(* Logix 5000 project; controller R400_500_XLS vendor 1 type 14 code 216 rev 31.11; software revision 31.01; part 17 of 32 *)
(* tags used below, declared in another part *)
   bResetAllCycle : BOOL;
   Calib : SINT;
   CalibCnt : SINT;   // Calibration Step Counter
   CalibData : UDT_SCALE[8];
   CalibEnabled : BOOL;   // RTD Calibration Enabled bit
   CalibIndex : DINT;   // Calibration Pointer
   CustomCycleIterator : DINT;
   CycleDryingStandard : UDT_DRY;
   CycleModifBuffer : UDT_CYCLE;
   Cycles : UDT_CYCLE[11];
   CyclesDefault : UDT_CYCLE[7];   // Preliminary Data block to reset Cycles Values
   CycleSmartDryingHeatSens : UDT_DRY;
   CycleSmartDryingRegular : UDT_DRY;
   CycleWith_NonRecircFRinseDefault : UDT_FRINSE;
   CycleWith_RecircFRinseDefault : UDT_FRINSE;
   CycleWithoutDry : UDT_DRY;
   CycleWithoutFRinseWithoutTankDefault : UDT_FRINSE;
   CycleWithoutFRinseWithTankDefault : UDT_FRINSE;
   DESCALER : SINT;
   DRYING : DINT;   // Drying id number
   ENVIRO_CARE : SINT;
   EXTRA_CARE : SINT;
   FC83_AutoSpeed : BOOL;   // Cycle pump speed selection
   FC83_AutoWtrLevel : BOOL;   // Cycle water level selection
   FC83_CyclePerm : BOOL;   // Cycle permission selection
   M : DINT[5];   // Memory Bits
   ONS_FC84 : SINT;
   PLASTIC_CARE : SINT;
   ResetCycleName : BOOL;
   RINSE_CARE : SINT;
   Run : DINT;
   STANDARD : SINT;
   Supervisor : DINT;
   USER_DEFINED_11 : SINT;
   USER_DEFINED_7 : SINT;
   CycleName : STRING[12];
   CycleNameDefault : STRING[12];
   CyclePtr : DINT;   // Cycle Pointeur
   DryTemp : REAL;
   I_Dry_RTD : DINT;   // Drying RTD
   I_Pw_Tnk_RTD : DINT;   // Pure water tank RTD
   I_Smp_RTD : DINT;   // Sump RTD
   NumInput : UDT_NUMERIC_INPUT[65];   // Numeric input
   PureWaterTankTemp : REAL;   // Pure water tank temperature
   Screen_Ctrl : DINT;   // PLC Screen Request
   StringInput : UDT_STRING_INPUT[6];
   SumpTemp : REAL;   // Sump temperature in °C
   Tpb : DINT[11];
   TpbImage : DINT[11];
   Unit : Hrdwre;   // Unit Configuration
(* MainProgram, continued *)

ROUTINE SPV_4_CycleNames   (* ladder *)
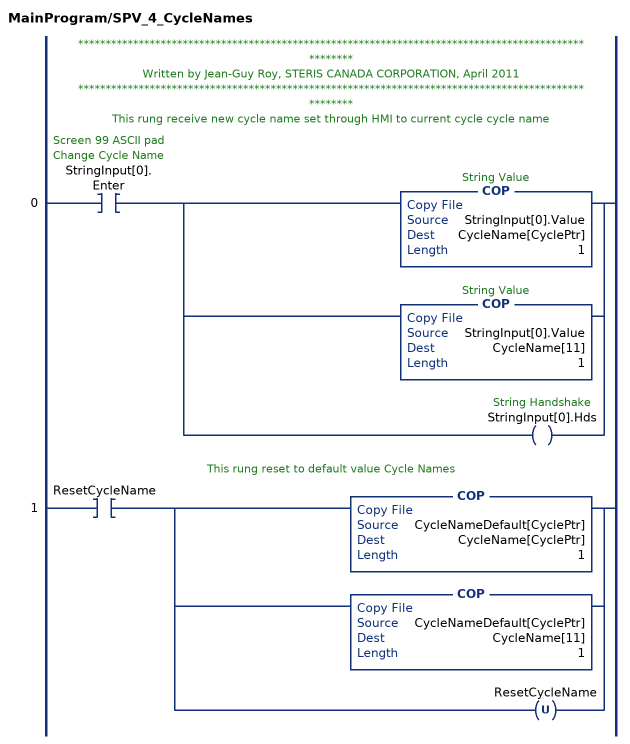
   // ****************************************************************************************************
   // Written by Jean-Guy Roy, STERIS CANADA CORPORATION, April 2011
   // ****************************************************************************************************
   // This rung receive new cycle name set through HMI to current cycle cycle name
   0: XIC(StringInput[0].Enter)[COP(StringInput[0].Value,CycleName[CyclePtr],1) ,COP(StringInput[0].Value,CycleName[11],1) ,OTE(StringInput[0].Hds) ];
   // This rung reset to default value Cycle Names
   1: XIC(ResetCycleName)[COP(CycleNameDefault[CyclePtr],CycleName[CyclePtr],1) ,COP(CycleNameDefault[CyclePtr],CycleName[11],1) ,OTU(ResetCycleName) ];
END_ROUTINE

ROUTINE SPV_8_ResetToDefaultCyclesValues   (* ladder *)
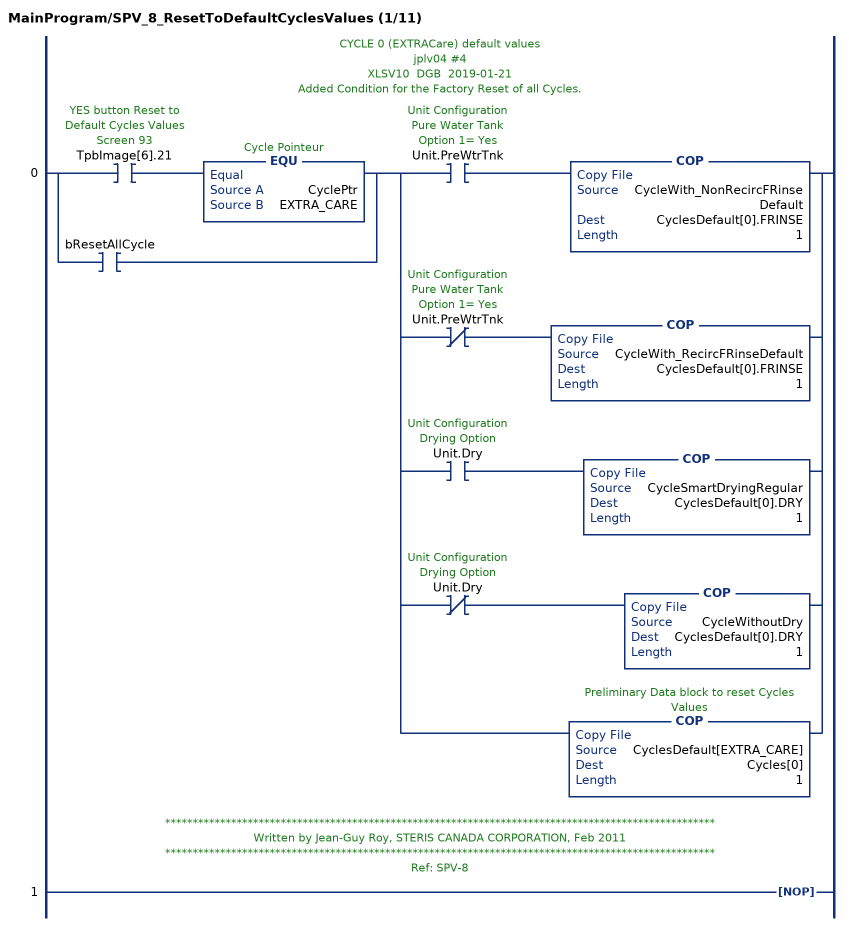
   // CYCLE 0 (EXTRACare) default values
   // jplv04 #4
   // XLSV10  DGB  2019-01-21
   // Added Condition for the Factory Reset of all Cycles.
   0: [XIC(TpbImage[6].21) EQU(CyclePtr,EXTRA_CARE) ,XIC(bResetAllCycle) ][XIC(Unit.PreWtrTnk) COP(CycleWith_NonRecircFRinseDefault,CyclesDefault[0].FRINSE,1) ,XIO(Unit.PreWtrTnk) COP(CycleWith_RecircFRinseDefault,CyclesDefault[0].FRINSE,1) ,XIC(Unit.Dry) COP(CycleSmartDryingRegular,CyclesDefault[0].DRY,1) ,XIO(Unit.Dry) COP(CycleWithoutDry,CyclesDefault[0].DRY,1) ,COP(CyclesDefault[EXTRA_CARE],Cycles[0],1) ];
   // ****************************************************************************************************
   // Written by Jean-Guy Roy, STERIS CANADA CORPORATION, Feb 2011
   // ****************************************************************************************************
   // Ref: SPV-8
   1: NOP();
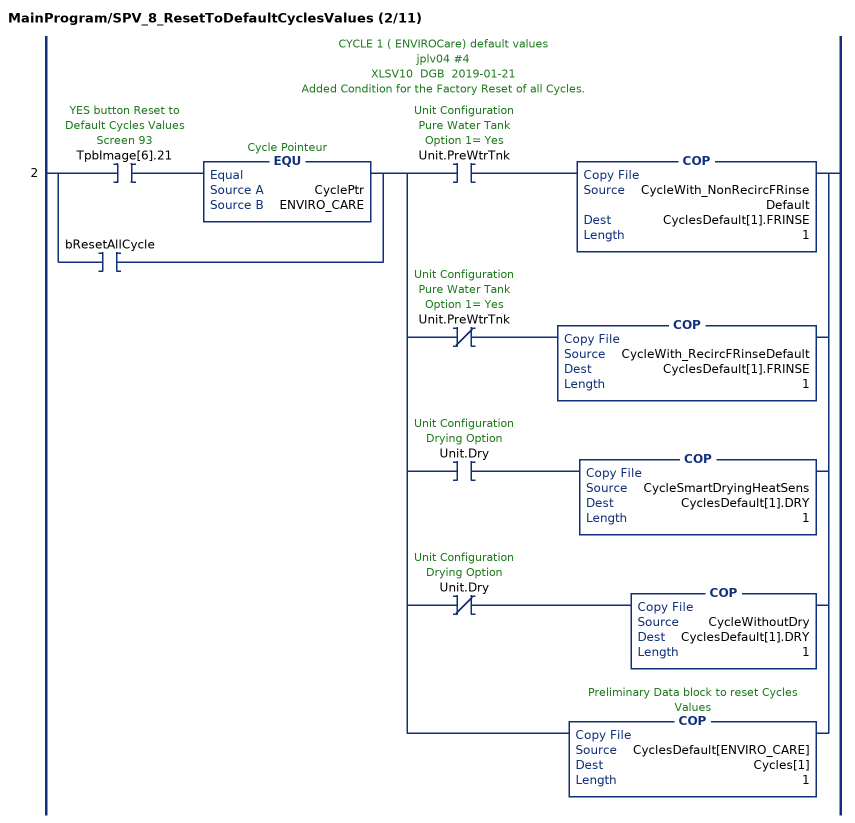
   // CYCLE 1 ( ENVIROCare) default values
   // jplv04 #4
   // XLSV10  DGB  2019-01-21
   // Added Condition for the Factory Reset of all Cycles.
   2: [XIC(TpbImage[6].21) EQU(CyclePtr,ENVIRO_CARE) ,XIC(bResetAllCycle) ][XIC(Unit.PreWtrTnk) COP(CycleWith_NonRecircFRinseDefault,CyclesDefault[1].FRINSE,1) ,XIO(Unit.PreWtrTnk) COP(CycleWith_RecircFRinseDefault,CyclesDefault[1].FRINSE,1) ,XIC(Unit.Dry) COP(CycleSmartDryingHeatSens,CyclesDefault[1].DRY,1) ,XIO(Unit.Dry) COP(CycleWithoutDry,CyclesDefault[1].DRY,1) ,COP(CyclesDefault[ENVIRO_CARE],Cycles[1],1) ];
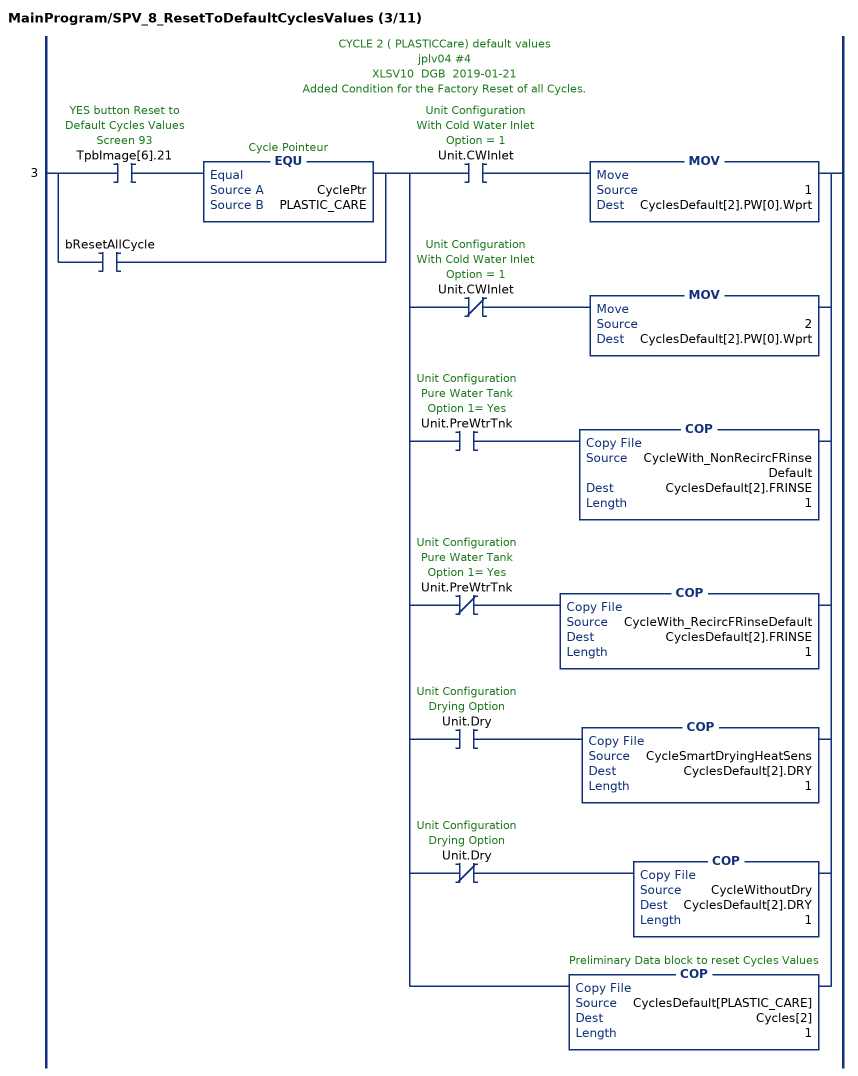
   // CYCLE 2 ( PLASTICCare) default values
   // jplv04 #4
   // XLSV10  DGB  2019-01-21
   // Added Condition for the Factory Reset of all Cycles.
   3: [XIC(TpbImage[6].21) EQU(CyclePtr,PLASTIC_CARE) ,XIC(bResetAllCycle) ][XIC(Unit.CWInlet) MOV(1,CyclesDefault[2].PW[0].Wprt) ,XIO(Unit.CWInlet) MOV(2,CyclesDefault[2].PW[0].Wprt) ,XIC(Unit.PreWtrTnk) COP(CycleWith_NonRecircFRinseDefault,CyclesDefault[2].FRINSE,1) ,XIO(Unit.PreWtrTnk) COP(CycleWith_RecircFRinseDefault,CyclesDefault[2].FRINSE,1) ,XIC(Unit.Dry) COP(CycleSmartDryingHeatSens,CyclesDefault[2].DRY,1) ,XIO(Unit.Dry) COP(CycleWithoutDry,CyclesDefault[2].DRY,1) ,COP(CyclesDefault[PLASTIC_CARE],Cycles[2],1) ];
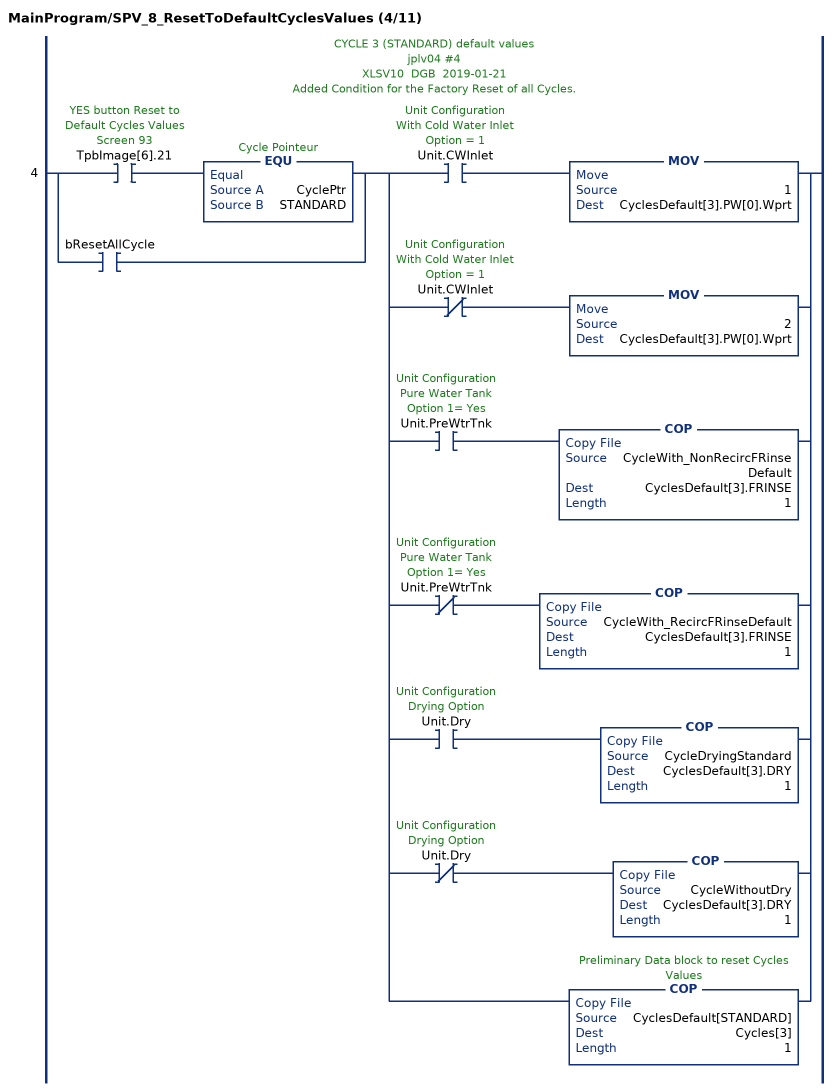
   // CYCLE 3 (STANDARD) default values
   // jplv04 #4
   // XLSV10  DGB  2019-01-21
   // Added Condition for the Factory Reset of all Cycles.
   4: [XIC(TpbImage[6].21) EQU(CyclePtr,STANDARD) ,XIC(bResetAllCycle) ][XIC(Unit.CWInlet) MOV(1,CyclesDefault[3].PW[0].Wprt) ,XIO(Unit.CWInlet) MOV(2,CyclesDefault[3].PW[0].Wprt) ,XIC(Unit.PreWtrTnk) COP(CycleWith_NonRecircFRinseDefault,CyclesDefault[3].FRINSE,1) ,XIO(Unit.PreWtrTnk) COP(CycleWith_RecircFRinseDefault,CyclesDefault[3].FRINSE,1) ,XIC(Unit.Dry) COP(CycleDryingStandard,CyclesDefault[3].DRY,1) ,XIO(Unit.Dry) COP(CycleWithoutDry,CyclesDefault[3].DRY,1) ,COP(CyclesDefault[STANDARD],Cycles[3],1) ];
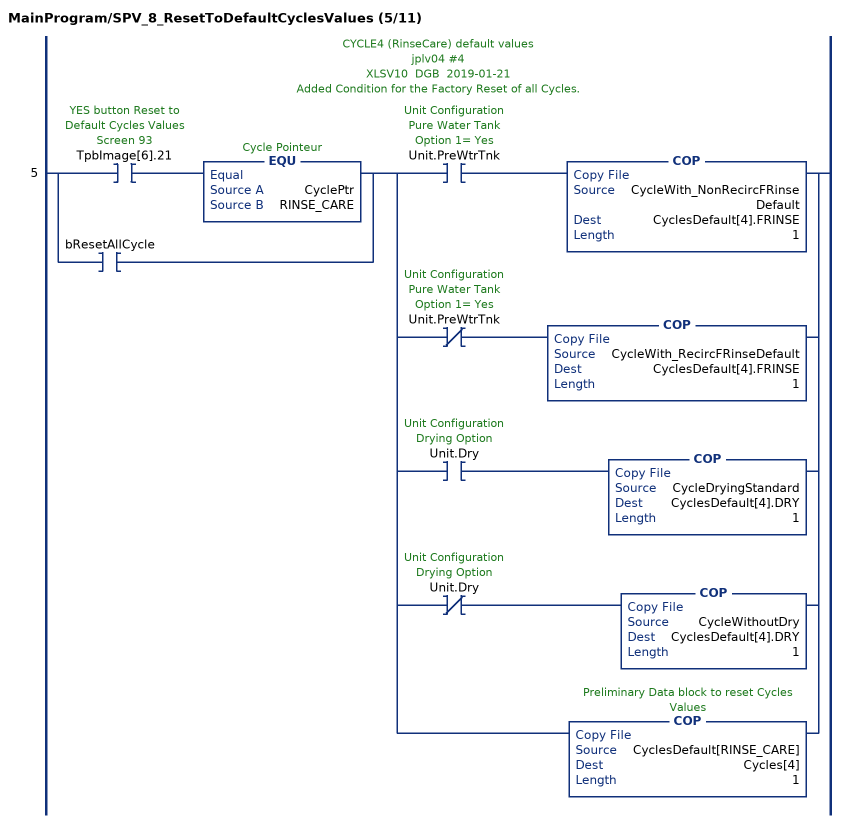
   // CYCLE4 (RinseCare) default values
   // jplv04 #4
   // XLSV10  DGB  2019-01-21
   // Added Condition for the Factory Reset of all Cycles.
   5: [XIC(TpbImage[6].21) EQU(CyclePtr,RINSE_CARE) ,XIC(bResetAllCycle) ][XIC(Unit.PreWtrTnk) COP(CycleWith_NonRecircFRinseDefault,CyclesDefault[4].FRINSE,1) ,XIO(Unit.PreWtrTnk) COP(CycleWith_RecircFRinseDefault,CyclesDefault[4].FRINSE,1) ,XIC(Unit.Dry) COP(CycleDryingStandard,CyclesDefault[4].DRY,1) ,XIO(Unit.Dry) COP(CycleWithoutDry,CyclesDefault[4].DRY,1) ,COP(CyclesDefault[RINSE_CARE],Cycles[4],1) ];
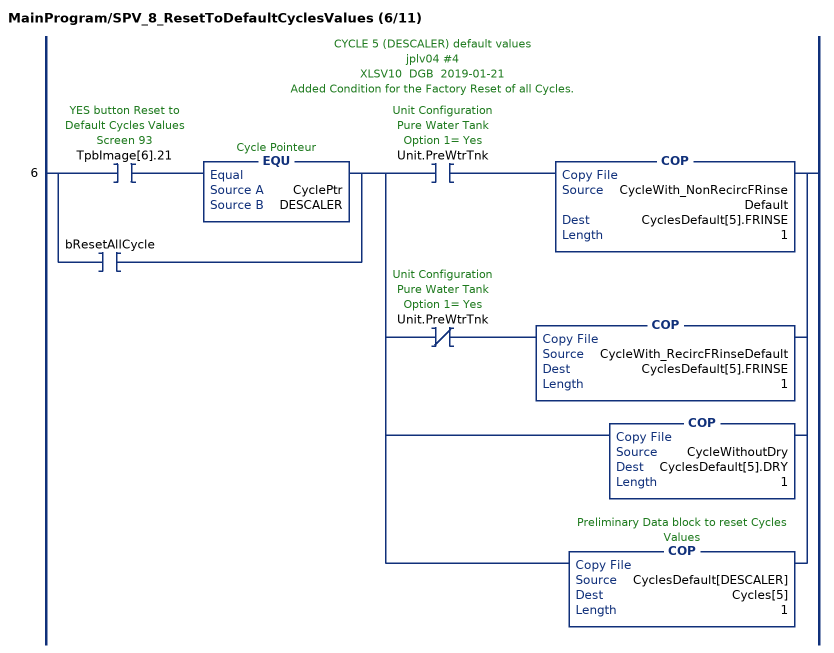
   // CYCLE 5 (DESCALER) default values
   // jplv04 #4
   // XLSV10  DGB  2019-01-21
   // Added Condition for the Factory Reset of all Cycles.
   6: [XIC(TpbImage[6].21) EQU(CyclePtr,DESCALER) ,XIC(bResetAllCycle) ][XIC(Unit.PreWtrTnk) COP(CycleWith_NonRecircFRinseDefault,CyclesDefault[5].FRINSE,1) ,XIO(Unit.PreWtrTnk) COP(CycleWith_RecircFRinseDefault,CyclesDefault[5].FRINSE,1) ,COP(CycleWithoutDry,CyclesDefault[5].DRY,1) ,COP(CyclesDefault[DESCALER],Cycles[5],1) ];
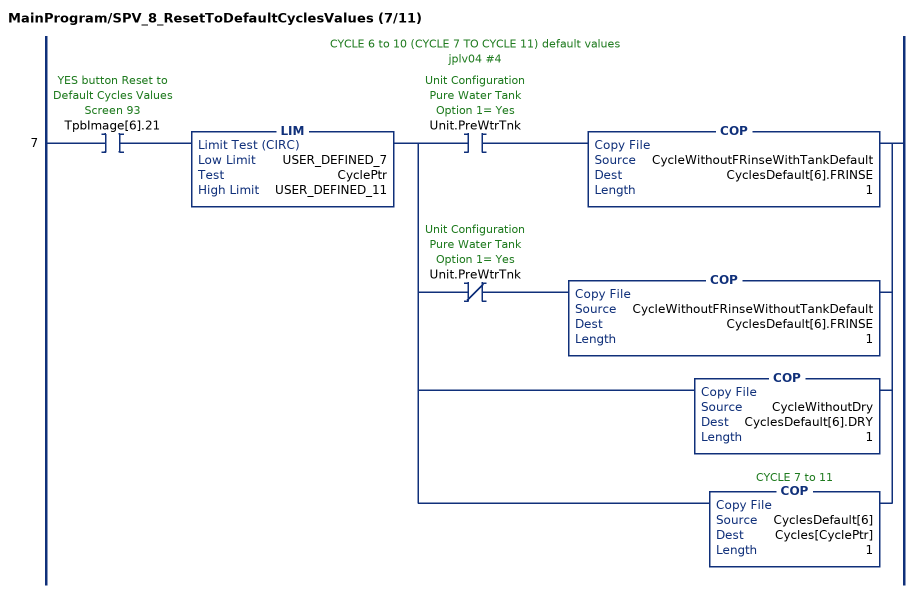
   // CYCLE 6 to 10 (CYCLE 7 TO CYCLE 11) default values
   // jplv04 #4
   7: XIC(TpbImage[6].21)LIM(USER_DEFINED_7,CyclePtr,USER_DEFINED_11)[XIC(Unit.PreWtrTnk) COP(CycleWithoutFRinseWithTankDefault,CyclesDefault[6].FRINSE,1) ,XIO(Unit.PreWtrTnk) COP(CycleWithoutFRinseWithoutTankDefault,CyclesDefault[6].FRINSE,1) ,COP(CycleWithoutDry,CyclesDefault[6].DRY,1) ,COP(CyclesDefault[6],Cycles[CyclePtr],1) ];
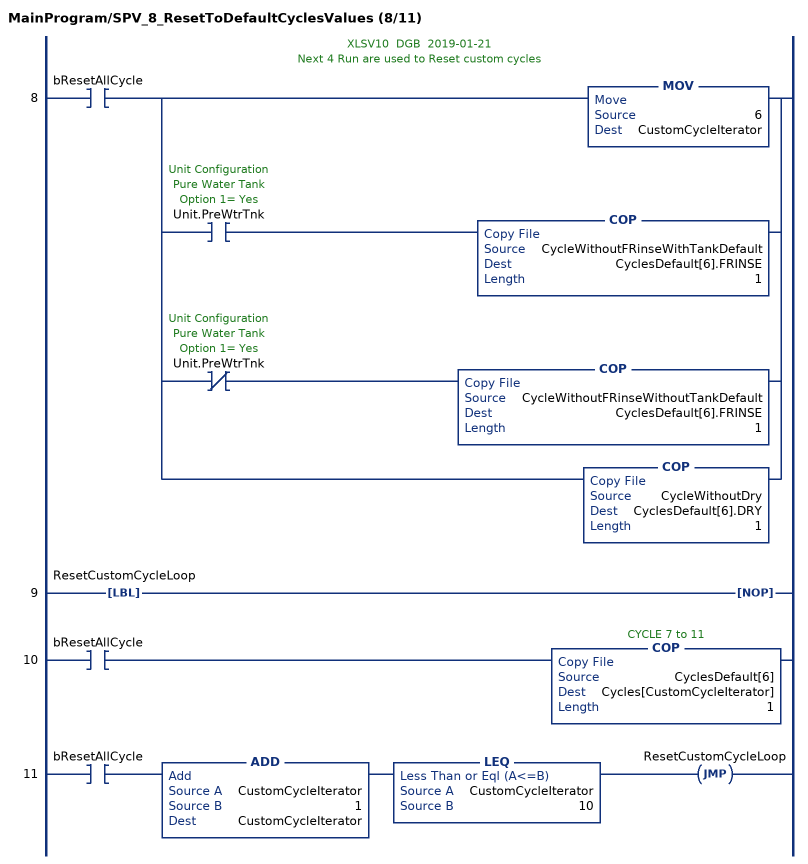
   // XLSV10  DGB  2019-01-21
   // Next 4 Run are used to Reset custom cycles
   8: XIC(bResetAllCycle)[MOV(6,CustomCycleIterator) ,XIC(Unit.PreWtrTnk) COP(CycleWithoutFRinseWithTankDefault,CyclesDefault[6].FRINSE,1) ,XIO(Unit.PreWtrTnk) COP(CycleWithoutFRinseWithoutTankDefault,CyclesDefault[6].FRINSE,1) ,COP(CycleWithoutDry,CyclesDefault[6].DRY,1) ];
   9: LBL(ResetCustomCycleLoop)NOP();
   10: XIC(bResetAllCycle)COP(CyclesDefault[6],Cycles[CustomCycleIterator],1);
   11: XIC(bResetAllCycle)ADD(CustomCycleIterator,1,CustomCycleIterator)LEQ(CustomCycleIterator,10)JMP(ResetCustomCycleLoop);
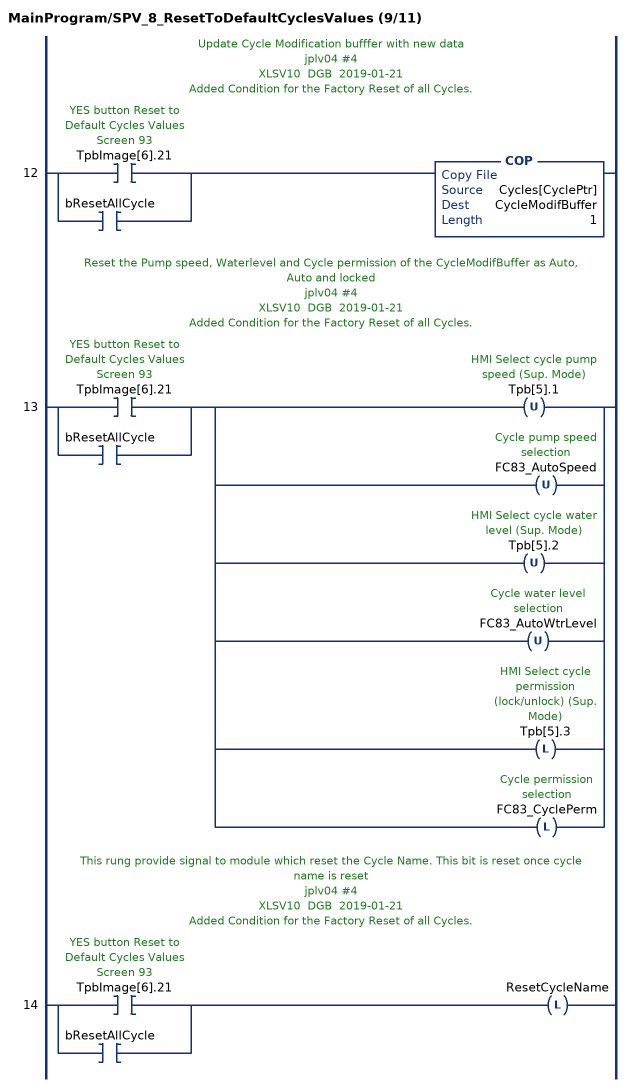
   // Update Cycle Modification bufffer with new data
   // jplv04 #4
   // XLSV10  DGB  2019-01-21
   // Added Condition for the Factory Reset of all Cycles.
   12: [XIC(TpbImage[6].21) ,XIC(bResetAllCycle) ]COP(Cycles[CyclePtr],CycleModifBuffer,1);
   // Reset the Pump speed, Waterlevel and Cycle permission of the CycleModifBuffer as Auto, Auto and locked
   // jplv04 #4
   // XLSV10  DGB  2019-01-21
   // Added Condition for the Factory Reset of all Cycles.
   13: [XIC(TpbImage[6].21) ,XIC(bResetAllCycle) ][OTU(Tpb[5].1) ,OTU(FC83_AutoSpeed) ,OTU(Tpb[5].2) ,OTU(FC83_AutoWtrLevel) ,OTL(Tpb[5].3) ,OTL(FC83_CyclePerm) ];
   // This rung provide signal to module which reset the Cycle Name. This bit is reset once cycle name is reset
   // jplv04 #4
   // XLSV10  DGB  2019-01-21
   // Added Condition for the Factory Reset of all Cycles.
   14: [XIC(TpbImage[6].21) ,XIC(bResetAllCycle) ]OTL(ResetCycleName);
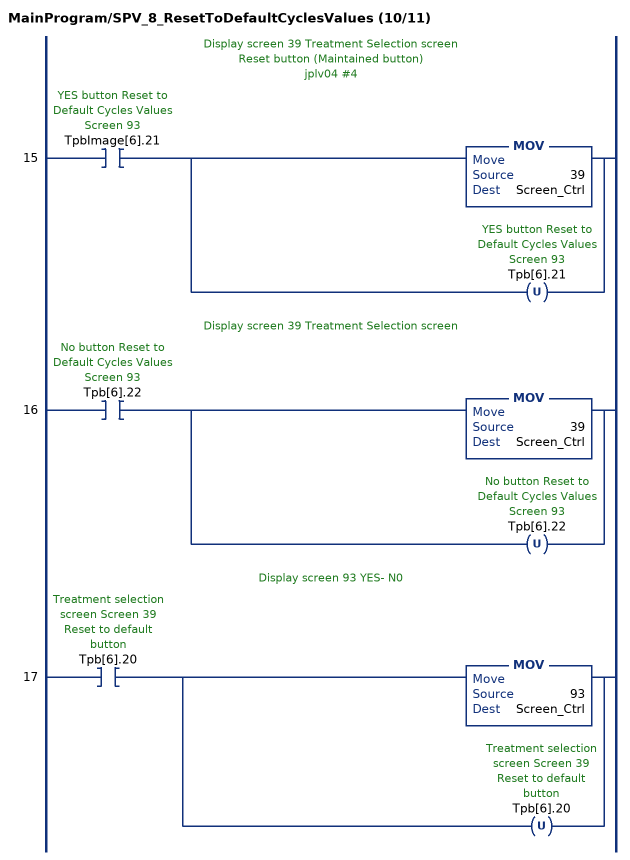
   // Display screen 39 Treatment Selection screen
   // Reset button (Maintained button)
   // jplv04 #4
   15: XIC(TpbImage[6].21)[MOV(39,Screen_Ctrl) ,OTU(Tpb[6].21) ];
   // Display screen 39 Treatment Selection screen
   16: XIC(Tpb[6].22)[MOV(39,Screen_Ctrl) ,OTU(Tpb[6].22) ];
   // Display screen 93 YES- N0
   17: XIC(Tpb[6].20)[MOV(93,Screen_Ctrl) ,OTU(Tpb[6].20) ];
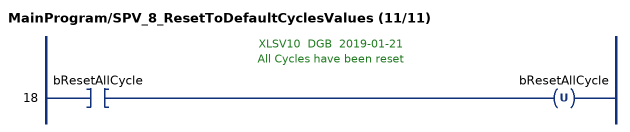
   // XLSV10  DGB  2019-01-21
   // All Cycles have been reset
   18: XIC(bResetAllCycle)OTU(bResetAllCycle);
END_ROUTINE

ROUTINE SPV_9_RTD_CALIBRATION   (* ladder *)
// Routine for the calibration of the analog inputs
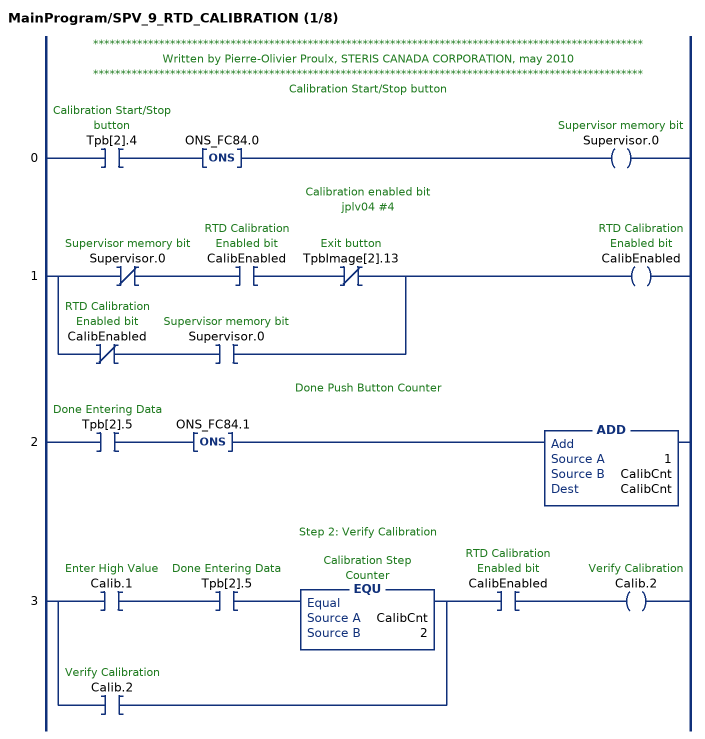
   // ****************************************************************************************************
   // Written by Pierre-Olivier Proulx, STERIS CANADA CORPORATION, may 2010
   // ****************************************************************************************************
   // Calibration Start/Stop button
   0: XIC(Tpb[2].4)ONS(ONS_FC84.0)OTE(Supervisor.0);
   // Calibration enabled bit
   // jplv04 #4
   1: [XIO(Supervisor.0) XIC(CalibEnabled) XIO(TpbImage[2].13) ,XIO(CalibEnabled) XIC(Supervisor.0) ]OTE(CalibEnabled);
   // Done Push Button Counter
   2: XIC(Tpb[2].5)ONS(ONS_FC84.1)ADD(1,CalibCnt,CalibCnt);
   // Step 2: Verify Calibration
   3: [XIC(Calib.1) XIC(Tpb[2].5) EQU(CalibCnt,2) ,XIC(Calib.2) ]XIC(CalibEnabled)OTE(Calib.2);
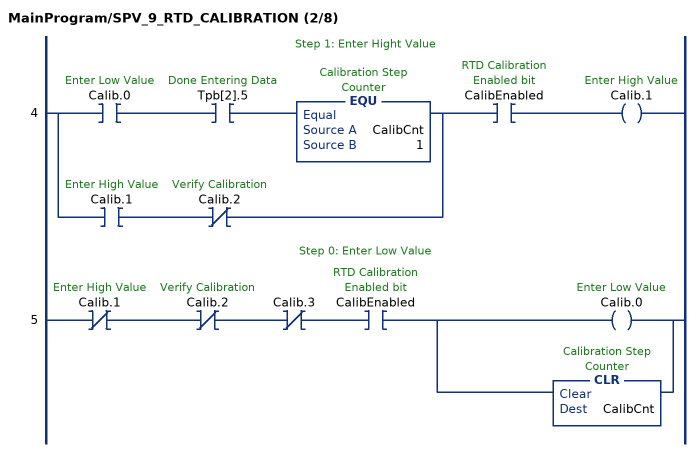
   // Step 1: Enter Hight Value
   4: [XIC(Calib.0) XIC(Tpb[2].5) EQU(CalibCnt,1) ,XIC(Calib.1) XIO(Calib.2) ]XIC(CalibEnabled)OTE(Calib.1);
   // Step 0: Enter Low Value
   5: XIO(Calib.1)XIO(Calib.2)XIO(Calib.3)XIC(CalibEnabled)[OTE(Calib.0) ,CLR(CalibCnt) ];
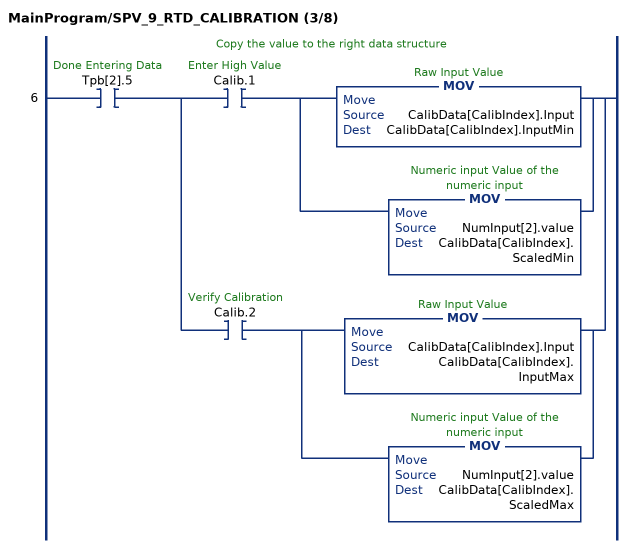
   // Copy the value to the right data structure
   6: XIC(Tpb[2].5)[XIC(Calib.1) [MOV(CalibData[CalibIndex].Input,CalibData[CalibIndex].InputMin) ,MOV(NumInput[2].value,CalibData[CalibIndex].ScaledMin) ] ,XIC(Calib.2) [MOV(CalibData[CalibIndex].Input,CalibData[CalibIndex].InputMax) ,MOV(NumInput[2].value,CalibData[CalibIndex].ScaledMax) ] ];
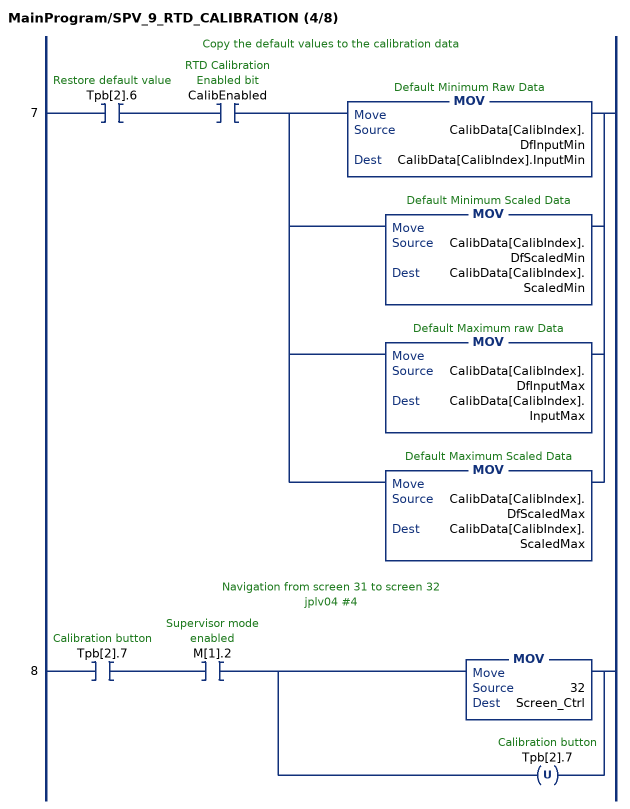
   // Copy the default values to the calibration data
   7: XIC(Tpb[2].6)XIC(CalibEnabled)[MOV(CalibData[CalibIndex].DfInputMin,CalibData[CalibIndex].InputMin) ,MOV(CalibData[CalibIndex].DfScaledMin,CalibData[CalibIndex].ScaledMin) ,MOV(CalibData[CalibIndex].DfInputMax,CalibData[CalibIndex].InputMax) ,MOV(CalibData[CalibIndex].DfScaledMax,CalibData[CalibIndex].ScaledMax) ];
   // Navigation from screen 31 to screen 32
   // jplv04 #4
   8: XIC(Tpb[2].7)XIC(M[1].2)[MOV(32,Screen_Ctrl) ,OTU(Tpb[2].7) ];
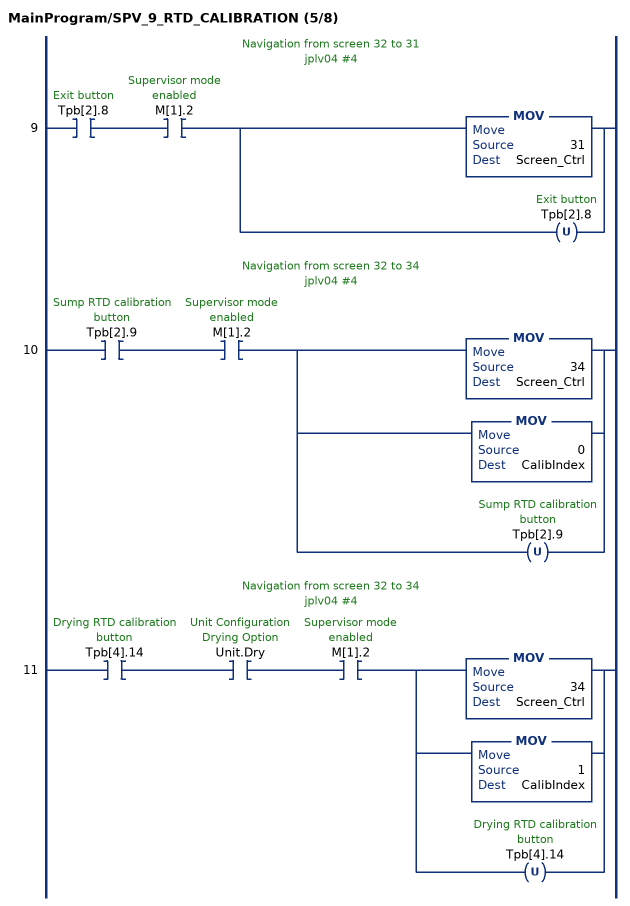
   // Navigation from screen 32 to 31
   // jplv04 #4
   9: XIC(Tpb[2].8)XIC(M[1].2)[MOV(31,Screen_Ctrl) ,OTU(Tpb[2].8) ];
   // Navigation from screen 32 to 34
   // jplv04 #4
   10: XIC(Tpb[2].9)XIC(M[1].2)[MOV(34,Screen_Ctrl) ,MOV(0,CalibIndex) ,OTU(Tpb[2].9) ];
   // Navigation from screen 32 to 34
   // jplv04 #4
   11: XIC(Tpb[4].14)XIC(Unit.Dry)XIC(M[1].2)[MOV(34,Screen_Ctrl) ,MOV(1,CalibIndex) ,OTU(Tpb[4].14) ];
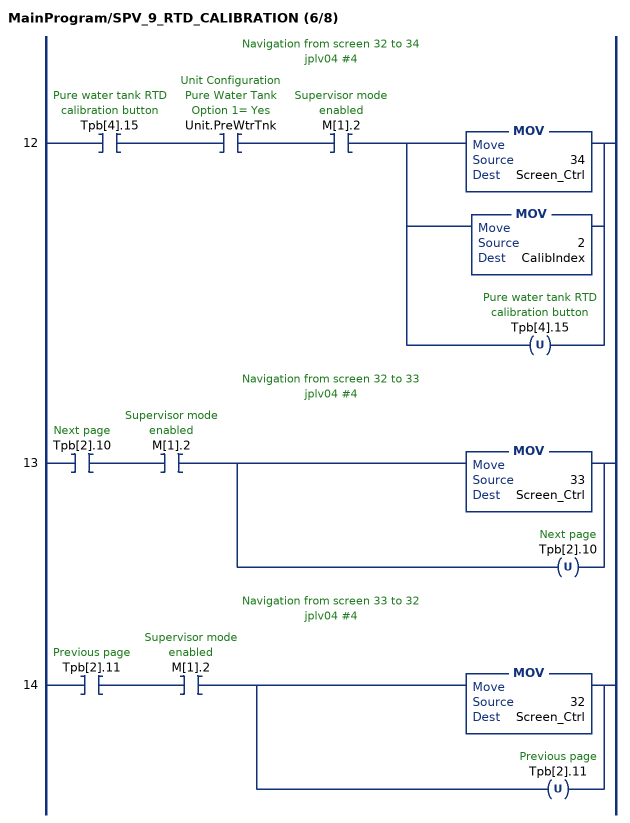
   // Navigation from screen 32 to 34
   // jplv04 #4
   12: XIC(Tpb[4].15)XIC(Unit.PreWtrTnk)XIC(M[1].2)[MOV(34,Screen_Ctrl) ,MOV(2,CalibIndex) ,OTU(Tpb[4].15) ];
   // Navigation from screen 32 to 33
   // jplv04 #4
   13: XIC(Tpb[2].10)XIC(M[1].2)[MOV(33,Screen_Ctrl) ,OTU(Tpb[2].10) ];
   // Navigation from screen 33 to 32
   // jplv04 #4
   14: XIC(Tpb[2].11)XIC(M[1].2)[MOV(32,Screen_Ctrl) ,OTU(Tpb[2].11) ];
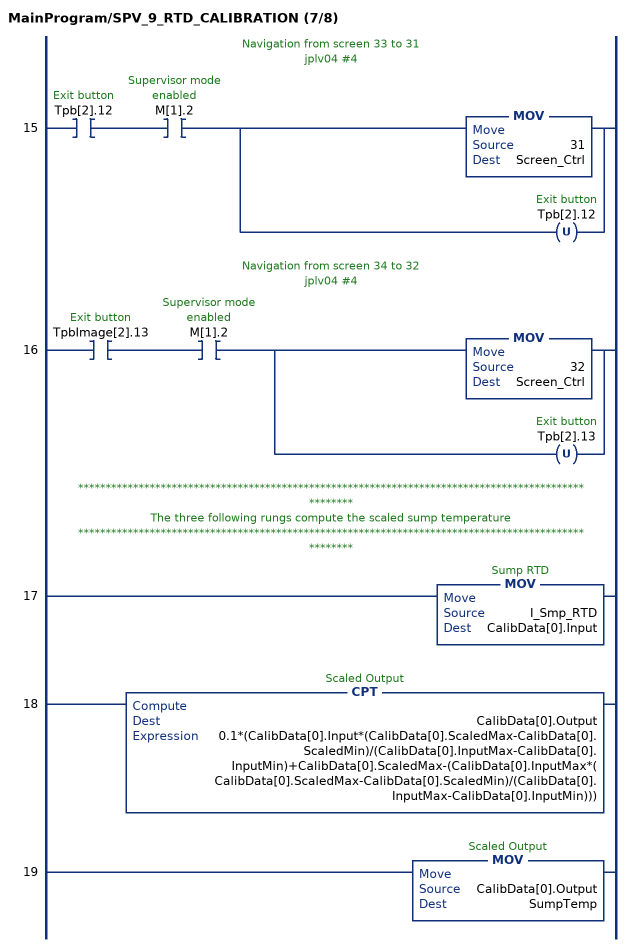
   // Navigation from screen 33 to 31
   // jplv04 #4
   15: XIC(Tpb[2].12)XIC(M[1].2)[MOV(31,Screen_Ctrl) ,OTU(Tpb[2].12) ];
   // Navigation from screen 34 to 32
   // jplv04 #4
   16: XIC(TpbImage[2].13)XIC(M[1].2)[MOV(32,Screen_Ctrl) ,OTU(Tpb[2].13) ];
   // ****************************************************************************************************
   // The three following rungs compute the scaled sump temperature
   // ****************************************************************************************************
   17: MOV(I_Smp_RTD,CalibData[0].Input);
   18: CPT(CalibData[0].Output,0.1*(CalibData[0].Input*(CalibData[0].ScaledMax-CalibData[0].ScaledMin)/(CalibData[0].InputMax-CalibData[0].InputMin)+CalibData[0].ScaledMax-(CalibData[0].InputMax*(CalibData[0].ScaledMax-CalibData[0].ScaledMin)/(CalibData[0].InputMax-CalibData[0].InputMin))));
   19: MOV(CalibData[0].Output,SumpTemp);
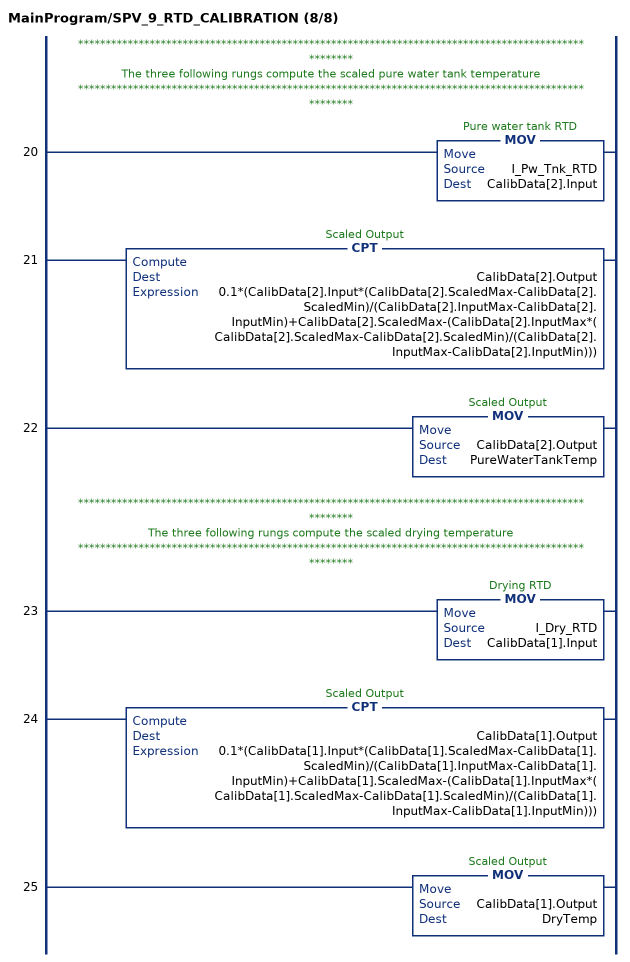
   // ****************************************************************************************************
   // The three following rungs compute the scaled pure water tank temperature
   // ****************************************************************************************************
   20: MOV(I_Pw_Tnk_RTD,CalibData[2].Input);
   21: CPT(CalibData[2].Output,0.1*(CalibData[2].Input*(CalibData[2].ScaledMax-CalibData[2].ScaledMin)/(CalibData[2].InputMax-CalibData[2].InputMin)+CalibData[2].ScaledMax-(CalibData[2].InputMax*(CalibData[2].ScaledMax-CalibData[2].ScaledMin)/(CalibData[2].InputMax-CalibData[2].InputMin))));
   22: MOV(CalibData[2].Output,PureWaterTankTemp);
   // ****************************************************************************************************
   // The three following rungs compute the scaled drying temperature
   // ****************************************************************************************************
   23: MOV(I_Dry_RTD,CalibData[1].Input);
   24: CPT(CalibData[1].Output,0.1*(CalibData[1].Input*(CalibData[1].ScaledMax-CalibData[1].ScaledMin)/(CalibData[1].InputMax-CalibData[1].InputMin)+CalibData[1].ScaledMax-(CalibData[1].InputMax*(CalibData[1].ScaledMax-CalibData[1].ScaledMin)/(CalibData[1].InputMax-CalibData[1].InputMin))));
   25: MOV(CalibData[1].Output,DryTemp);
END_ROUTINE
